Fanuc KAREL source: ko00049.KL

-- PROVISIONAL review KL for V1013-1; original PC SHA256 828da7a068ef2bc1be8602638f045d11819ff7d843c51241d2a380c9e066ef53
-- Incomplete behavior may be omitted. Consult companion uncertainty JSON. Do not deploy.
PROGRAM KO00049
%NOLOCKGROUP
BEGIN
  -- UNRESOLVED_PC offsets 5-12; opcodes 9D,23
  -- UNRESOLVED_PC offsets 17-66; opcodes 27,27,49,7E,AD,22,1C,22,31,7E,4A
  -- UNRESOLVED_PC offsets 71-75; opcodes 7F
END KO00049
